Universal Robots URScript: T007_curved_weld_hybrid.urscript

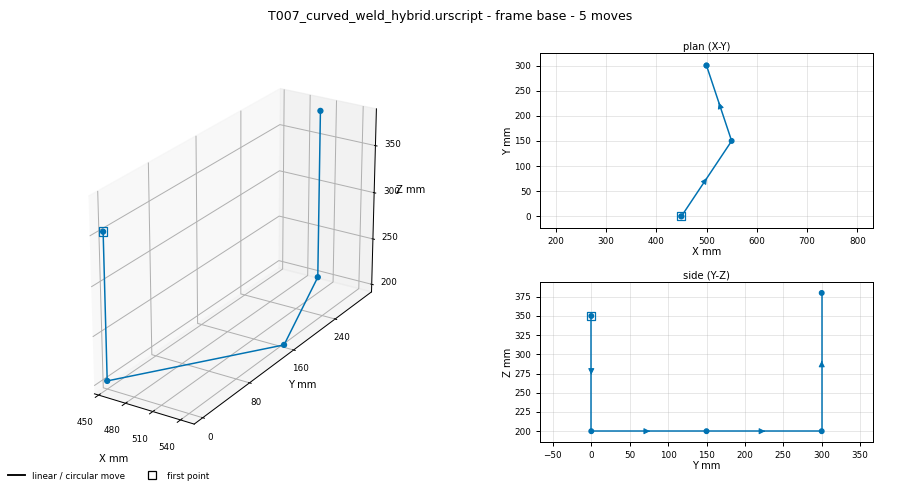
[picture p0: tool path of T007_curved_weld_hybrid.urscript in frame base, 5 of 7 moves have a stored position in this frame; points joined in program order, loops and branches not executed]
# Task: T007 — Curved contour weld — hybrid mode
# Generated by ENFIELD IR→URScript Translator
# Operating mode: hybrid | Max TCP speed: 0.300 m/s
# Robot: ur5e
#
# WARNING: This is auto-generated code for SIMULATION ONLY.
# Do NOT deploy to a physical robot without safety review.

def task_T007():
  # Safety preamble: tool centre point and payload declared before motion
  set_tcp(p[0.0000, 0.0000, 0.1600, 0.0, 0.0, 0.0])
  set_payload(3.500)

  # [0] Verify E-Stop clear
  # E-Stop safety check (hardware-enforced on UR controller)
  if (get_digital_in(0) == True):
    popup("E-Stop active — aborting program.", error=True)
    halt
  end

  # [1] Home position
  movej([0.0000, -1.5708, 1.5708, -1.5708, -1.5708, 0.0000], a=1.4000, v=0.7500)

  # [2] Approach above weld fixture
  movel(p[0.450000, 0.000000, 0.350000, 0.0000, 3.1416, 0.0000], a=1.0000, v=0.2500, r=0.0100)

  # [3] Descend to weld start
  movel(p[0.450000, 0.000000, 0.200000, 0.0000, 3.1416, 0.0000], a=0.5000, v=0.1000, r=0.0010)

  # [4] Gas pre-flow ON
  set_digital_out(1, True)

  # [5] Gas stabilization
  sleep(0.5000)

  # [6] Arc ON
  # Welding arc ON (I=150A, wire=6.0m/min)
  set_digital_out(0, True)   # arc enable
  set_analog_out(0, 0.500)  # current (normalized)
  set_analog_out(1, 0.400)  # wire feed (normalized)

  # [7] Weld midpoint
  movel(p[0.550000, 0.150000, 0.200000, 0.0000, 3.1416, 0.0000], a=0.2000, v=0.0600, r=0.0050)

  # [8] Weld end
  movel(p[0.500000, 0.300000, 0.200000, 0.0000, 3.1416, 0.0000], a=0.2000, v=0.0600)

  # [9] Arc OFF
  # Welding arc OFF
  set_digital_out(0, False)
  set_analog_out(0, 0.0)
  set_analog_out(1, 0.0)

  # [10] Post-weld gas flow
  sleep(1.0000)

  # [11] Gas flow OFF
  set_digital_out(1, False)

  # [12] Retract above weld end
  movel(p[0.500000, 0.300000, 0.380000, 0.0000, 3.1416, 0.0000], a=1.0000, v=0.2500, r=0.0100)

  # [13] Return to home
  movej([0.0000, -1.5708, 1.5708, -1.5708, -1.5708, 0.0000], a=1.4000, v=0.7500)

end

# Entry point
task_T007()
